Fanuc KAREL source: KO00027.KL

PROGRAM KO00027
%NOLOCKGROUP
VAR
  P1: JOINTPOS
  P2: JOINTPOS
  P3: JOINTPOS
  OUT: XYZWPREXT
BEGIN
  OUT = FRAME(P1, P2, P3)
END KO00027
